SUBAPPLICATION Button_IXA_TO_logiBUS_QXA_BG_OPC (* Button IXA -> logiBUS QXA + Hintergrundfarbe, plus OPC-UA Read/Write (generisch, ein Kanal) *)
  (* Standard: 61499-2; Description: Copyright (c) 2023 Meisterschulen am Ostbahnhof This program and the accompanying materials are made available under the terms of the Eclipse Public License 2.0 which is available at https://www.eclipse.org/legal/epl-2.0/ SPDX-License-Identifier: EPL-2.0 *)
  (* Version 1.3, 2026-11-06, Franz Höpfinger, Meisterschulen am Ostbahnhof, AX_OR_2 durch AX_LAST_2 ersetzt (last writer wins): mit READ und WRITE auf demselben Knoten hielt das Echo des eigenen PUBLISH den Ausgang ueber das ODER dauerhaft EIN *)
  (* Version 1.2, 2026-09-07, Franz Höpfinger, Meisterschulen am Ostbahnhof, Vorruebergehend non-latching: SR-Latch (AX_ASR_RF_TRIG x2 + ASR_MERGE_2 + ASR_AX_SR) durch einfaches AX_OR_2 ersetzt - Button UND Remote-Kommando sind jetzt tastend (Pegel), kein Klick-Toggle mehr *)
  (* Version 1.1, 2026-07-20, Franz Höpfinger, Meisterschulen am Ostbahnhof, Background *)
  (* Version 1.0, 2026-01-15, Franz Höpfinger, Meisterschulen am Ostbahnhof, initial API and implementation and/or initial documentation *)
  PACKAGE MyLib::sys;
  IMPORT isobus::UT::Q::const::IDs::ID_NULL;
  IMPORT logiBUS::io::DQ::logiBUS_DO;
  IMPORT logiBUS::io::DQ::logiBUS_DO_S;
  (* Documentation:
  Button → logiBUS-Ausgang (wer zuletzt schreibt, gewinnt)
   Lokaler VT-Button und Remote-OPC-UA-Kommando laufen über AX_LAST_2: Die Quelle, die zuletzt einen Wert geliefert hat, bestimmt den Ausgang. Der Ausgang wird per PUBLISH auf ID_WRITE gemeldet.
   Liegen ID_READ und ID_WRITE auf demselben Knoten, kommt das eigene PUBLISH als SUBSCRIBE zurück. Mit dem früheren AX_OR_2 blieb der Ausgang dadurch dauerhaft EIN. Mit AX_LAST_2 ist das Echo gleich dem aktuellen Wert und ändert nichts.
   Für die vorherige Klick-Toggle-Variante (SR-Latch, ein Klick EIN, nächster Klick AUS) Button_IXA_TO_logiBUS_QXA_BG_OPC_LATCHING verwenden - identisches Interface, 1:1 austauschbar.
  *)
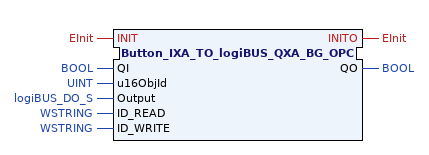
  EVENT_INPUT
    INIT : EInit; (* Initialization Request *)
  END_EVENT
  EVENT_OUTPUT
    INITO : EInit; (* Initialization Confirm *)
  END_EVENT
  VAR_INPUT
    QI : BOOL := TRUE; (* Quality Input - TRUE to enable service *)
    u16ObjId : UINT := ID_NULL; (* Object ID Button/Hintergrund (VT), ID_NULL = noch kein VT-Objekt *)
    Output : logiBUS::io::DQ::logiBUS_DO_S := logiBUS_DO::Invalid; (* Identify the Output Output_Q1..Q12 *)
    ID_READ : WSTRING; (* OPC-UA Subscribe-Key (schreibbar) *)
    ID_WRITE : WSTRING; (* OPC-UA Publish-Key (lesbar) *)
  END_VAR
  VAR_OUTPUT
    QO : BOOL; (* Quality Output - TRUE if service executed successfully *)
  END_VAR
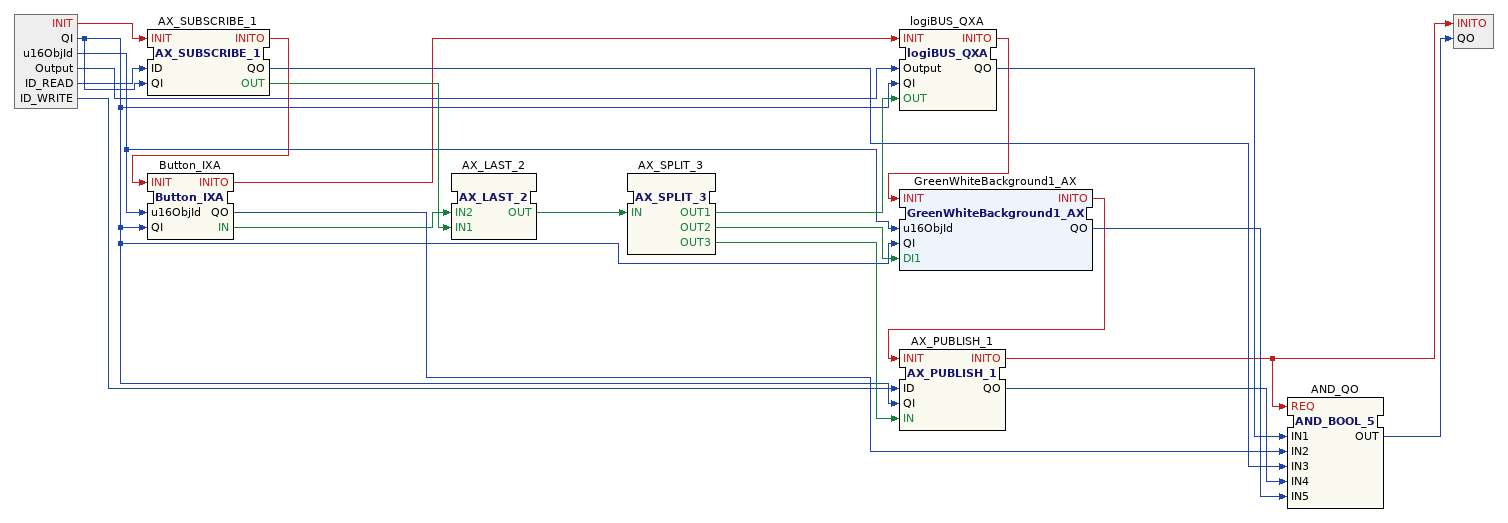
  FBS
    logiBUS_QXA : logiBUS::io::DQ::logiBUS_QXA;
    Button_IXA : isobus::UT::io::Button::Button_IXA;
    AX_SUBSCRIBE_1 : adapter::net::AX_SUBSCRIBE_1;
    AX_PUBLISH_1 : adapter::net::AX_PUBLISH_1;
    AX_LAST_2 : adapter::events::unidirectional::AX_LAST_2;
    AX_SPLIT_3 : adapter::events::unidirectional::AX_SPLIT_3;
    AND_QO : iec61131::booleanOperators::AND_BOOL_5;
  END_FBS
  SUBAPPS
    GreenWhiteBackground1_AX : MyLib::sys::GreenWhiteBackground1_AX;
  END_SUBAPPS
  EVENT_CONNECTIONS
    INIT TO AX_SUBSCRIBE_1.INIT;
    AX_SUBSCRIBE_1.INITO TO Button_IXA.INIT;
    Button_IXA.INITO TO logiBUS_QXA.INIT;
    GreenWhiteBackground1_AX.INITO TO AX_PUBLISH_1.INIT;
    logiBUS_QXA.INITO TO GreenWhiteBackground1_AX.INIT;
    AX_PUBLISH_1.INITO TO AND_QO.REQ;
    AX_PUBLISH_1.INITO TO INITO;
  END_CONNECTIONS
  DATA_CONNECTIONS
    u16ObjId TO Button_IXA.u16ObjId;
    Output TO logiBUS_QXA.Output;
    u16ObjId TO GreenWhiteBackground1_AX.u16ObjId;
    ID_READ TO AX_SUBSCRIBE_1.ID;
    ID_WRITE TO AX_PUBLISH_1.ID;
    QI TO logiBUS_QXA.QI;
    QI TO Button_IXA.QI;
    QI TO AX_SUBSCRIBE_1.QI;
    QI TO AX_PUBLISH_1.QI;
    logiBUS_QXA.QO TO AND_QO.IN1;
    Button_IXA.QO TO AND_QO.IN2;
    AX_SUBSCRIBE_1.QO TO AND_QO.IN3;
    AX_PUBLISH_1.QO TO AND_QO.IN4;
    AND_QO.OUT TO QO;
    QI TO GreenWhiteBackground1_AX.QI;
    GreenWhiteBackground1_AX.QO TO AND_QO.IN5;
  END_CONNECTIONS
  ADAPTER_CONNECTIONS
    Button_IXA.IN TO AX_LAST_2.IN2;
    AX_SUBSCRIBE_1.OUT TO AX_LAST_2.IN1;
    AX_SPLIT_3.OUT1 TO logiBUS_QXA.OUT;
    AX_SPLIT_3.OUT2 TO GreenWhiteBackground1_AX.DI1;
    AX_SPLIT_3.OUT3 TO AX_PUBLISH_1.IN;
    AX_LAST_2.OUT TO AX_SPLIT_3.IN;
  END_CONNECTIONS
END_SUBAPPLICATION
